// TIA Portal V19 export
TYPE "EM03_Output"
   STRUCT
      Status : "EM_Output";
      FeedActive : Bool;   // AlimentaciÃ³n/agua en regulaciÃ³n
      LevelInterlock : Bool;   // Nivel mÃ­nimo no permitido: regulaciÃ³n bloqueada
   END_STRUCT;
END_TYPE
